FUNCTION_BLOCK "Q12"
VERSION : 0.1

VAR_INPUT
    THICKNESS_FAULT : BOOL;
    THICKNESS_SIGNAL_VALID : BOOL;
    CUTTING_RUN : BOOL;
    FaultTimestamp : DINT;
    CycleTime : TIME := T#10ms;
END_VAR

VAR_OUTPUT
    THICKNESS_ALARM : BOOL;
    Slab_Fault_Counter : UINT;
    Slab_Runtime_Accumulator : LTIME;
    Slab_Fault_History : ARRAY[0..4] OF DINT;
END_VAR

VAR
    PreviousValidFault : BOOL := FALSE;
    HoldElapsed : LTIME := LTIME#0ns;
    HoldActive : BOOL := FALSE;
    HistoryFilled : INT := 0;
    ShiftIndex : INT := 0;
    CycleNs : LTIME := LTIME#0ns;
END_VAR

BEGIN
    // Elapsed interval represented by this invocation, expressed in nanoseconds.
    CycleNs := DINT_TO_LTIME(TIME_TO_DINT(CycleTime) * 1000);

    IF NOT THICKNESS_SIGNAL_VALID THEN
        // Signal lost: alarm off, holding state cleared, no logging and no runtime accrual.
        THICKNESS_ALARM := FALSE;
        HoldActive := FALSE;
        HoldElapsed := LTIME#0ns;
        PreviousValidFault := FALSE;
    ELSE
        IF HoldActive THEN
            HoldElapsed := HoldElapsed + CycleNs;
            IF HoldElapsed >= DINT_TO_LTIME(500000000) THEN
                HoldActive := FALSE;
                HoldElapsed := LTIME#0ns;
            END_IF;
        END_IF;

        IF THICKNESS_FAULT AND (NOT PreviousValidFault) THEN
            // New valid thickness fault: count it and store the newest timestamp.
            IF Slab_Fault_Counter < 65535 THEN
                Slab_Fault_Counter := Slab_Fault_Counter + 1;
            END_IF;

            IF HistoryFilled < 5 THEN
                FOR ShiftIndex := HistoryFilled TO 1 BY -1 DO
                    Slab_Fault_History[ShiftIndex] := Slab_Fault_History[ShiftIndex - 1];
                END_FOR;
                Slab_Fault_History[0] := FaultTimestamp;
                HistoryFilled := HistoryFilled + 1;
            ELSE
                FOR ShiftIndex := 4 TO 1 BY -1 DO
                    Slab_Fault_History[ShiftIndex] := Slab_Fault_History[ShiftIndex - 1];
                END_FOR;
                Slab_Fault_History[0] := FaultTimestamp;
            END_IF;

            HoldActive := TRUE;
            HoldElapsed := LTIME#0ns;
        END_IF;

        PreviousValidFault := THICKNESS_FAULT;

        IF THICKNESS_FAULT OR HoldActive THEN
            THICKNESS_ALARM := TRUE;
        ELSE
            THICKNESS_ALARM := FALSE;
        END_IF;

        IF CUTTING_RUN AND (NOT THICKNESS_FAULT) THEN
            Slab_Runtime_Accumulator := Slab_Runtime_Accumulator + CycleNs;
        END_IF;
    END_IF;
END_FUNCTION_BLOCK
